(* IEC 61131-3 sources: generating_plc_code_with_llms/Code#1/Platypus2/second run, 5 files *)

(* ---- 12.st ---- *)
// 9.104289531707764s
// 1
function sinh(x)
    return exp(x)*cosh(x);
end_function

(* ---- 11.st ---- *)
// 61.69238305091858s
// 1
program main;

// Declare variables and constants
integer i, n;
real x;
constant pi = 3.14159265358979323846264338327950288419716939937510;

// Function definition
function sign(x)
    input real x;
    output integer s;

    if (x > 0.0) then
        s := 1;
    elseif (x < 0.0) then
        s := -1;
    else
        s := 0;
    end_if;
end_function;

// Main program logic
write("Enter a number: ");
read(n);

write("The sign of ", n, " is ", sign(n));

stop;

(* ---- 13.st ---- *)
// 19.646280527114868s
// 2
REPEAT
    IF (SELECTED_NUMBER = 10) THEN
        EXIT
    END_IF
END_REPEAT

(* ---- 15.st ---- *)
// 30.642439126968384s
// 2
IF (E_A = 0) THEN
    IF (P_HU = 0 AND P_AL = 1) THEN
        P_AL = 0
    END_IF
END_IF

(* ---- 19.st ---- *)
// 68.69949984550476s
// 2
```
THICKNESS(MD_1)
D_MAX := MD_1;
D_MIN := MD_1;
IF (S1 = 0) THEN
    IF (D_MAX > V_MAX OR D_MIN < V_MIN) THEN
        P1 := TRUE;
    ELSE
        P1 := FALSE;
    END_IF;
END_IF;
```
